(* PLC project Unnamed, Unknown Unnamed 1 *)
(* stored: creationDateTime 2026-11-17T11:02:30, modificationDateTime 2026-11-17T15:16:27 *)

PROGRAM Main
  VAR
    Button AT %IX0.0 : BOOL;
  END_VAR
  VAR
    Statelight : BOOL := TRUE;
  END_VAR
  VAR
    LEDG AT %QX0.0 : BOOL;
    LEDB AT %QX0.1 : BOOL;
    LEDR AT %QX0.2 : BOOL;
    LEDGu AT %QX0.3 : BOOL;
  END_VAR
  VAR
    TON0 : TON;
    OnTime : TIME := T#10s;
    OldState : BOOL;
    ButtonTimerState : BOOL := FALSE;
    TON1 : TON;
    ButtonTimer : TIME := T#80s;
    ButtonState : BOOL := FALSE;
    ButtonLightState : BOOL := FALSE;
    TON2 : TON;
    TON3 : TON;
  END_VAR

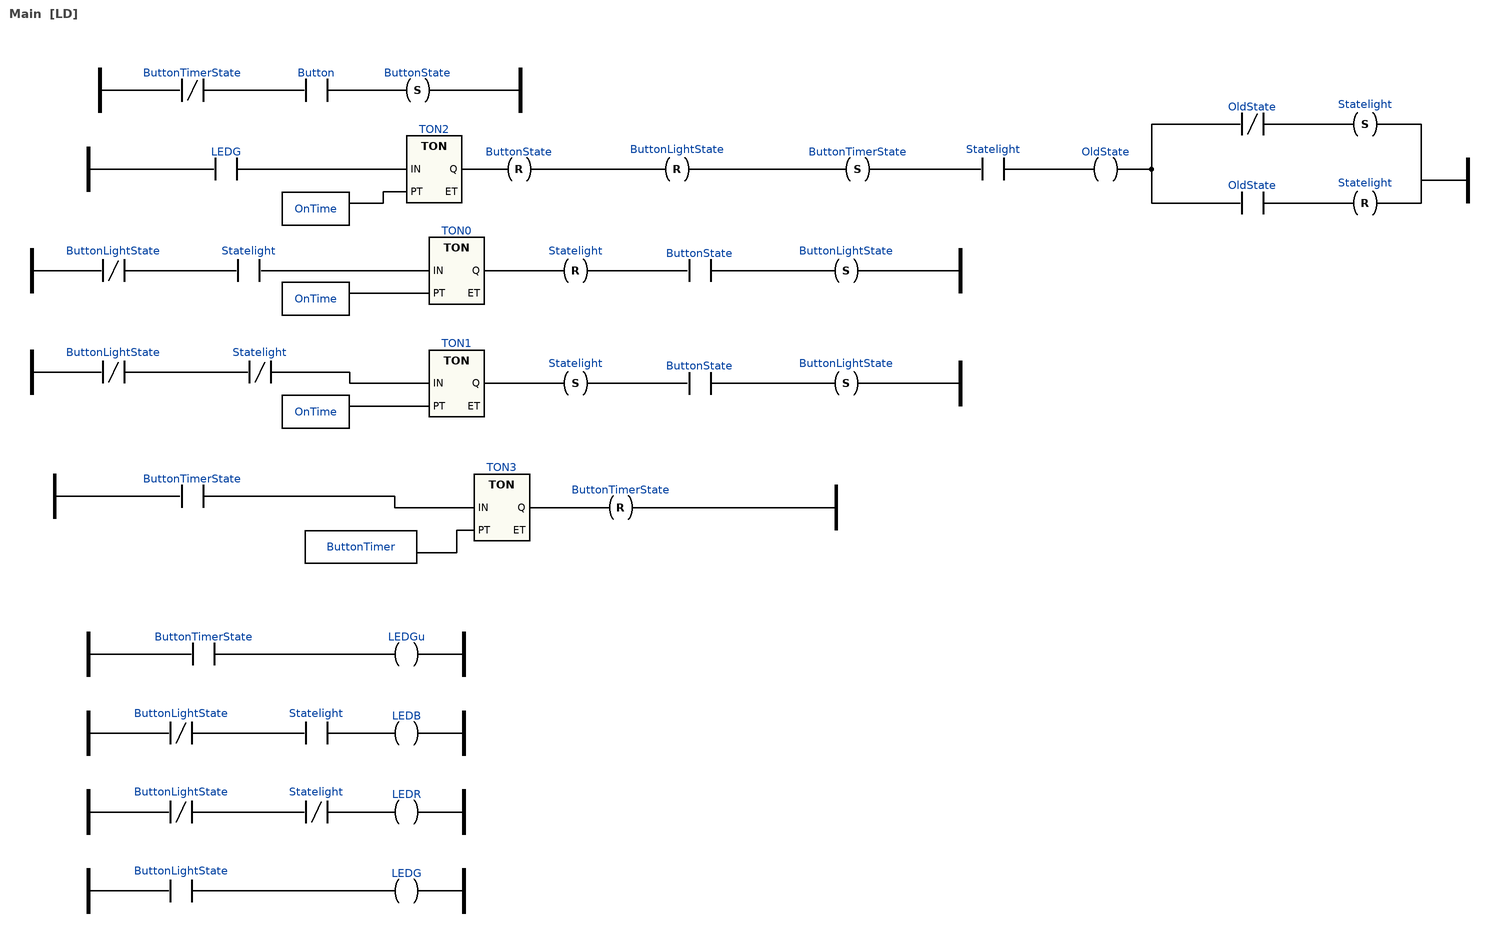
(* LD diagram, written out as Structured Text *)
LEDB := NOT ButtonLightState AND Statelight;
LEDR := NOT ButtonLightState AND NOT Statelight;
TON0(IN := NOT ButtonLightState AND Statelight, PT := OnTime);
IF TON0.Q THEN Statelight := FALSE; END_IF;
TON1(IN := NOT ButtonLightState AND NOT Statelight, PT := OnTime);
IF TON1.Q THEN Statelight := TRUE; END_IF;
IF NOT ButtonTimerState AND Button THEN ButtonState := TRUE; END_IF;
LEDG := ButtonLightState;
TON2(IN := LEDG, PT := OnTime);
IF TON2.Q THEN ButtonState := FALSE; END_IF;
IF TON2.Q THEN ButtonLightState := FALSE; END_IF;
IF TON0.Q AND ButtonState THEN ButtonLightState := TRUE; END_IF;
IF TON1.Q AND ButtonState THEN ButtonLightState := TRUE; END_IF;
IF TON2.Q AND Statelight AND NOT OldState THEN Statelight := TRUE; END_IF;
IF TON2.Q AND Statelight AND OldState THEN Statelight := FALSE; END_IF;
OldState := TON2.Q AND Statelight;
TON3(IN := ButtonTimerState, PT := ButtonTimer);
IF TON3.Q THEN ButtonTimerState := FALSE; END_IF;
IF TON2.Q THEN ButtonTimerState := TRUE; END_IF;
LEDGu := ButtonTimerState;
END_PROGRAM

CONFIGURATION Config0
  RESOURCE Res0 ON PLC
    TASK MainTask(INTERVAL := T#20ms, PRIORITY := 0);
    PROGRAM MainInstance WITH MainTask : Main;
  END_RESOURCE
END_CONFIGURATION
